(* IEC 61131-3 sources: iec-checker/test/st, 17 files *)

(* ---- declaration-analysis.st ---- *)
(* This demo includes some declaration errors *)
TYPE
    (* String types *)
    ST0 : STRING[5];                               (* OK *)
    ST1 : STRING;                                  (* OK *)
    ST2 : STRING[5] := 'foo';                      (* OK *)
    ST3 : STRING := 'platform_dependent';          (* OK *)
    ST4 : STRING[5] := "foobar";                   (* Error *)

    (* Subrange types *)
    ANALOG_DATA1 : INT (-4095 .. 4095);          (* OK *)
    ANALOG_DATA1 : INT (-4095 .. 4095) := 2000;  (* OK *)
    ANALOG_DATA1 : INT (-4095 .. 4095) := 4095;  (* OK: See 6.4.4.4.1 *)
    ANALOG_DATA1 : INT (-4095 .. 4095) := -4095; (* OK: See 6.4.4.4.1 *)
    ANALOG_DATA2 : INT (-4095 .. 4095) := 4099;  (* Error *)
    ANALOG_DATA2 : INT (-4095 .. 4095) := -4096; (* Error *)
END_TYPE

(* ---- merge-1.st ---- *)
TYPE example_struct :
  STRUCT
    Field : BOOL;
  END_STRUCT
END_TYPE

(* ---- plcopen-cp13.st ---- *)
(* Uncompatible: Recursive functions are forbidden *)
FUNCTION Factorial : INT
    VAR_INPUT
        X : INT;
    END_VAR

    IF X > 1 THEN
        Factorial := Factorial(X - 1) * X;
    ELSE
        Factorial := X;
    END_IF;
END_FUNCTION

(* Compatible iterative implementation *)
FUNCTION Factorial_good : INT
    VAR_INPUT
        X : INT;
    END_VAR
    VAR
        Acc : INT;
    END_VAR

    FOR I := 0 TO 100 DO
        Acc := Acc * X;
    END_FOR;
    Factorial := Acc;
END_FUNCTION

(* ---- plcopen-cp3.st ---- *)
FUNCTION demo : INT
    VAR_INPUT
        x1 : INT := 0;
        x2 : INT; (* PLCOPEN-CP3 *)
        x3 : STRING[5]; (* PLCOPEN-CP3 *)
        x4 : WSTRING[25] := 'spaces_disallowed';
        x5 : ARRAY [1..2, 1..3] OF INT; (* PLCOPEN-CP3 *)
        x6: ARRAY [0..7] OF BOOL := [0,1,1,0,0,1,0,0];
        x7 AT %B0 : INT;
    END_VAR
    x1 := 42;
END_FUNCTION

(* ---- plcopen-cp4.st ---- *)
FUNCTION demo : INT
    VAR_INPUT
        x1 AT %MX40 : INT; (* PLCOPEN-CP4 *)
        x2 AT %MX41 : INT; (* PLCOPEN-CP4 *)
        x3 AT %MX510 : INT;
    END_VAR
    x1 := 42;
END_FUNCTION

(* ---- plcopen-cp6.st ---- *)
FUNCTION demo : INT
    VAR_EXTERNAL
        x1 : INT; (* PLCOPEN-CP6 *)
    END_VAR
    x1 := 42;
END_FUNCTION

FUNCTION_BLOCK demo
    VAR_EXTERNAL
        x1 : INT; (* PLCOPEN-CP6 *)
    END_VAR
    x1 := 42;
END_FUNCTION_BLOCK

PROGRAM demo
    VAR_EXTERNAL
        x1 : INT;
    END_VAR
    x1 := 42;
END_PROGRAM

CLASS test1
  VAR_EXTERNAL
    x1 : INT;
  END_VAR

  METHOD PRIVATE count
    x1 := 42;
  END_METHOD

END_CLASS

(* ---- plcopen-cp9.st ---- *)
(* Example from PLCOpen guidelines, page 60.

   The following Function block CHARCURVE has:
   Number of Statements 18
   McCabe complexity of 12
   Prater complexity of 3,89
   Halstead complexity of 44,9
   Elshof complexity of 0,14

  NOTE: I'm not sure how they evaluated number of statements and appropriate
  complexity metrics. I have 4 additional statements for this program, and it
  seems correct for me.
 *)

FUNCTION_BLOCK CHARCURVE
  VAR_INPUT
    IN:INT;
    N:BYTE;
  END_VAR
  (* VAR_IN_OUT *)
    (* P : ARRAY [0 .. 10] OF POINT; *)
  (* END_VAR *)
  VAR_OUTPUT
    OUT:INT;
    ERR: BYTE;
  END_VAR
  VAR
    I:INT;
  END_VAR

  IF N > 1 AND N < 12 THEN
    ERR:=0;
    (* IF IN < P[0].X THEN *)
    IF IN < a THEN
      ERR := 2;
      OUT := DINT_TO_INT(a);
    (* ELSIF IN > P[N-1].X THEN *)
    ELSIF IN > a THEN
      ERR := 2;
      OUT := DINT_TO_INT(a);
    ELSE
      FOR I:=1 TO N-1 DO
        (* IF P[I-1].X >= P[I].X THEN *)
        IF a >= a THEN
          ERR:=1;
          EXIT;
        END_IF;
        (* IF IN <= P[I].X THEN *)
        IF IN <= a THEN
          EXIT;
        END_IF;
      END_FOR;
      IF ERR = 0 THEN
        (* OUT := DINT_TO_INT(P[I].Y - (P[I].X-IN) * (P[I].Y-P[I-1].Y) / (P[I].X-P[I-1].X)); *)
        OUT := DINT_TO_INT(a - (a - IN) * (a - a) / (a - a));
      ELSE
        OUT:=0;
      END_IF;
    END_IF;
  ELSE
    ERR := 4;
  END_IF;
END_FUNCTION_BLOCK

(* ---- dead-code.st ---- *)
FUNCTION dead_code_after_return : INT
  VAR
    counter : INT := 0;
    some_var : INT;
  END_VAR
  counter := counter + 1;
  counter := 2 + 2;
  RETURN;
  some_var := SQRT(16#42); (* UnreachableCode error *)
  some_var := 16#42; (* No additional warnings *)
  some_var := 19;
END_FUNCTION

PROGRAM dead_code_in_the_loops
VAR a : INT; i : INT; END_VAR
  WHILE i < 10 DO
    IF i = 5 THEN
      i := i + 1;
      EXIT;
      i := 19; (* UnreachableCode error *)
      i := 42; (* No additional warnings *)
      i := 42;
    ELSIF i = 6 THEN
      CONTINUE;
      i := 3; (* UnreachableCode error *)
      i := 44; (* No additional warnings *)
      i := 19;
    END_IF;
    i := i + 2;
  END_WHILE;
  I := 0;
END_PROGRAM

(* ---- merge-2.st ---- *)
PROGRAM Program1
  VAR
    instance AT %MW500 : example_struct;
  END_VAR

  %MW500 := TRUE;
END_PROGRAM

(* ---- plcopen-cp1.st ---- *)
(** PLCOPEN-CP1 – Access to a member shall be by name *)

PROGRAM program0
  VAR
    head AT %B0 : INT;
  END_VAR
  %B0 := 42;
END_PROGRAM

(* ---- plcopen-cp25.st ---- *)
PROGRAM demo
    VAR
        I : INT := 10;
        J : REAL := 0.55;
        a1 : BOOL; a2 : BYTE; a3 : WORD; a4 : DWORD; a5 : LWORD;
        b1 : SINT; b2 : INT; b3 : DINT; b4 : LINT;
        c1 : USINT; c2 : UINT; c3 : UDINT; c4 : ULINT;
        d1 : REAL; d2 : LREAL;
        e1 : TIME; e2 : LTIME;
        f1 : DT; f2 : LDT;
        g1 : DATE; g2 : LDATE;
        h1 : TOD; h2 : LTOD;
        i1 : CHAR; i2 : WCHAR; i3 : STRING[10]; i4 : WSTRING[10];
    END_VAR

  (* allowed implicit conversions *)
  a2 := a1; (* BOOL -> BYTE *)
  a3 := a2; (* BYTE -> WORD *)
  a4 := a3; (* WORD -> DWORD *)
  a5 := a4; (* DWORD -> LWORD *)

  b2 := b1; (* SINT -> INT *)
  b3 := b2; (* INT -> DINT *)
  b4 := b3; (* DINT -> LINT *)

  d2 := d1; (* REAL -> LREAL *)

  c2 := c1; (* USINT -> UINT *)
  c3 := c2; (* UINT -> UDINT *)
  c4 := c3; (* UDINT -> ULINT *)

  e2 := e1; (* TIME -> LTIME *)
  f2 := f1; (* DT -> LDT *)
  g2 := g1; (* DATE -> LDATE *)
  h2 := h1; (* TOD -> LTOD *)

  i2 := i1; (* CHAR -> WCHAR *)
  i4 := i3; (* STRING -> WSTRING *)

  i3 := i1; (* CHAR -> STRING *)
  i4 := i2; (* WCHAR -> WSTRING *)

  (* Implicit conversion not allowed - triggers warning *)
  I := J; (* REAL -> INT - not allowed *)

  (* Other examples of disallowed conversions *)
  b1 := b3; (* DINT -> SINT - not allowed *)
  c1 := c2; (* UINT -> USINT - not allowed *)
  a1 := a2; (* BYTE -> BOOL - not allowed *)
  d1 := d2; (* LREAL -> REAL - not allowed *)

  (* The correct way to write requires explicit conversion *)
  I := REAL_TO_INT(J);
  J := INT_TO_REAL(I);
  b1 := DINT_TO_SINT(b3);
  c1 := UINT_TO_USINT(c2);
  a1 := BYTE_TO_BOOL(a2);
  d1 := LREAL_TO_REAL(d2);

END_PROGRAM

(* ---- plcopen-cp28.st ---- *)
PROGRAM demo
    VAR
        x : TIME;
        y : TIME;
    END_VAR

    IF x = T#100MS THEN (* PLCOPEN CP-28 *)
      x := x + 1;
    END_IF;

    IF x <> T#100MS THEN (* PLCOPEN CP-28 *)
      x := x + 1;
    END_IF;

    IF T#100MS = x THEN (* PLCOPEN CP-28 *)
      x := x + 1;
    END_IF;

    IF T#100MS <> x THEN (* PLCOPEN CP-28 *)
      x := x + 1;
    END_IF;

    IF REAL_TO_INT(x) <> 0 THEN
      x := x + 1;
    END_IF;

    IF x >= T#100MS THEN
      x := x + 1;
    END_IF;

    IF x = y THEN
      x := x + 1;
    END_IF;
END_PROGRAM

(* ---- plcopen-cp8.st ---- *)
PROGRAM demo
    VAR
        x : REAL;
    END_VAR

    IF x = 0.0 THEN (* PLCOPEN CP-8 *)
      x := x + 1;
    END_IF;

    IF x <> 0.0 THEN (* PLCOPEN CP-8 *)
      x := x + 1;
    END_IF;

    IF 0.0 = x THEN (* PLCOPEN CP-8 *)
      x := x + 1;
    END_IF;

    IF 0.0 <> x THEN (* PLCOPEN CP-8 *)
      x := x + 1;
    END_IF;

    IF REAL_TO_INT(x) <> 0 THEN
      x := x + 1;
    END_IF;
END_PROGRAM

(* ---- plcopen-l10.st ---- *)
PROGRAM l10
  VAR
    i : INT := 0;
    j : INT := 0;
    flag : INT := 1;
    counter : INT := 0;
  END_VAR

  FOR i := 0 TO 10 DO
    FOR j := 10 TO 100 BY 2 DO
      IF flag THEN
        EXIT; (* PLCOPEN-CP10 *)
      END_IF;
      counter := counter + 1;
      IF j = 10 THEN
        CONTINUE; (* PLCOPEN-CP10 *)
      END_IF;
      EXIT; (* PLCOPEN-CP10 *)
    END_FOR;
  END_FOR;
END_PROGRAM

(* ---- plcopen-l17.st ---- *)
(** PLCOPEN-L17 – Each IF instruction should have an ELSE clause

    Reference: PLCopen Coding Guidelines 6.5.9. *)

PROGRAM program0
  VAR
    a : INT;
  END_VAR

  IF (a = 42) (* PLCOPEN-L17 *)
    THEN
      a := 0;
  END_IF;

  IF (a = 42) (* no warning *)
    THEN
      a := 0;
    ELSE
      a := 19;
  END_IF;

END_PROGRAM

(* ---- plcopen-n3.st ---- *)
PROGRAM program0
  VAR
    FOR_B : INT; (* PLCOPEN-N3 *)
    NO_FALSE_POSITIVE : INT;
    IF_A : INT; (* PLCOPEN-N3 *)
    TOF : INT; (* PLCOPEN-N3 *)
    OK_ALLOWED : INT;
  END_VAR

  FOR_B := IF_A / 1;
END_PROGRAM

(* ---- zero-division.st ---- *)
PROGRAM program0
  VAR_ACCESS
    acc : Var1 : DINT;
    acc : Var2 : DINT;
  END_VAR

  Var1 := 19 / 0;
  Var2 := Var1 / 1;
  Var2 := Var2 / 0;
END_PROGRAM
